SUBAPPLICATION TimedFunc (* Subapplication Type *)
  (* Standard: 61499-2 *)
  (* Version 1.0, 2023-01-29, Franz *)
  IMPORT isobus::UT::io::Softkey::SoftKeyActivationCode::SK_RELEASED;
  IMPORT isobus::UT::io::Auxiliary::IN::AuxiliaryState::AuxDisabled;
  IMPORT DataPanel::io::MI::DQ::DataPanel_MI_DO::Invalid;
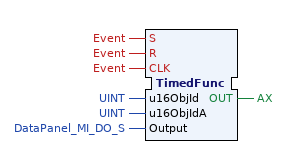
  EVENT_INPUT
    S; (* Set output Q *)
    R; (* Reset output Q *)
    CLK; (* Clock for triggering a output toggle *)
  END_EVENT
  VAR_INPUT
    u16ObjId : UINT;
    u16ObjIdA : UINT;
    Output : DataPanel::io::MI::DQ::DataPanel_MI_DO_S := Invalid;
  END_VAR
  PLUGS
    OUT : adapter::types::unidirectional::AX;
  END_PLUGS
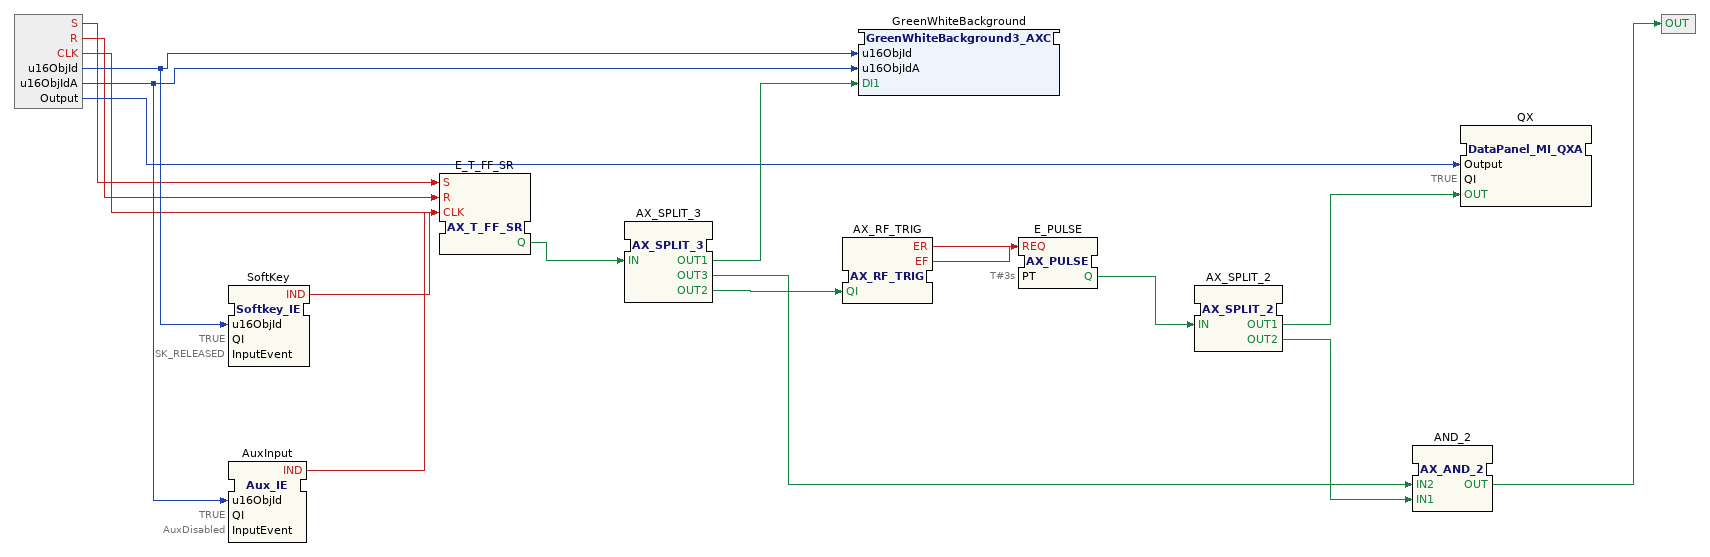
  FBS
    AND_2 : adapter::booleanOperators::AX_AND_2;
    QX : DataPanel::io::MI::DQ::DataPanel_MI_QXA(QI := TRUE);
    E_PULSE : adapter::events::unidirectional::timers::AX_PULSE(PT := T#3s);
    E_T_FF_SR : adapter::events::unidirectional::AX_T_FF_SR;
    AX_SPLIT_3 : adapter::events::unidirectional::AX_SPLIT_3;
    AX_RF_TRIG : adapter::events::unidirectional::AX_RF_TRIG;
    AX_SPLIT_2 : adapter::events::unidirectional::AX_SPLIT_2;
    SoftKey : isobus::UT::io::Softkey::Softkey_IE(QI := TRUE, InputEvent := SK_RELEASED);
    AuxInput : isobus::UT::io::Auxiliary::IN::Aux_IE(QI := TRUE, InputEvent := AuxDisabled);
  END_FBS
  SUBAPPS
    GreenWhiteBackground : MyLib::sys::GreenWhiteBackground3_AXC;
  END_SUBAPPS
  EVENT_CONNECTIONS
    S TO E_T_FF_SR.S;
    R TO E_T_FF_SR.R;
    CLK TO E_T_FF_SR.CLK;
    SoftKey.IND TO E_T_FF_SR.CLK;
    AuxInput.IND TO E_T_FF_SR.CLK;
    AX_RF_TRIG.ER TO E_PULSE.REQ;
    AX_RF_TRIG.EF TO E_PULSE.REQ;
  END_CONNECTIONS
  DATA_CONNECTIONS
    Output TO QX.Output;
    u16ObjIdA TO AuxInput.u16ObjId;
    u16ObjId TO SoftKey.u16ObjId;
    u16ObjId TO GreenWhiteBackground.u16ObjId;
    u16ObjIdA TO GreenWhiteBackground.u16ObjIdA;
  END_CONNECTIONS
  ADAPTER_CONNECTIONS
    E_T_FF_SR.Q TO AX_SPLIT_3.IN;
    AX_SPLIT_3.OUT1 TO GreenWhiteBackground.DI1;
    AX_SPLIT_3.OUT3 TO AND_2.IN2;
    E_PULSE.Q TO AX_SPLIT_2.IN;
    AX_SPLIT_2.OUT1 TO QX.OUT;
    AX_SPLIT_2.OUT2 TO AND_2.IN1;
    AND_2.OUT TO OUT;
    AX_SPLIT_3.OUT2 TO AX_RF_TRIG.QI;
  END_CONNECTIONS
END_SUBAPPLICATION
